Staubli VAL3: stop.pgx

program stop()
// Lab2A Level 3 - shared manual simulation / physical cycle
begin

  // Stop motion and feeding; preserve suction.
  resetMotion()

  trolleyOn = false
  barrierClosed = true
  blowOn = false

  if physicalRun
    taskKill("physicalIO")
    io:bOut2 = false
    io:bOut1 = false
    io:bOut5 = false
  endIf

  cycleStep = -1
  putln("Application stopped safely.")
  resetMotion()

end
